(* CODESYS project YarnStorage.xml

Project tree, tasks and I/O mapping:
  visualisation YarnStorage
*)

// /YarnStorage
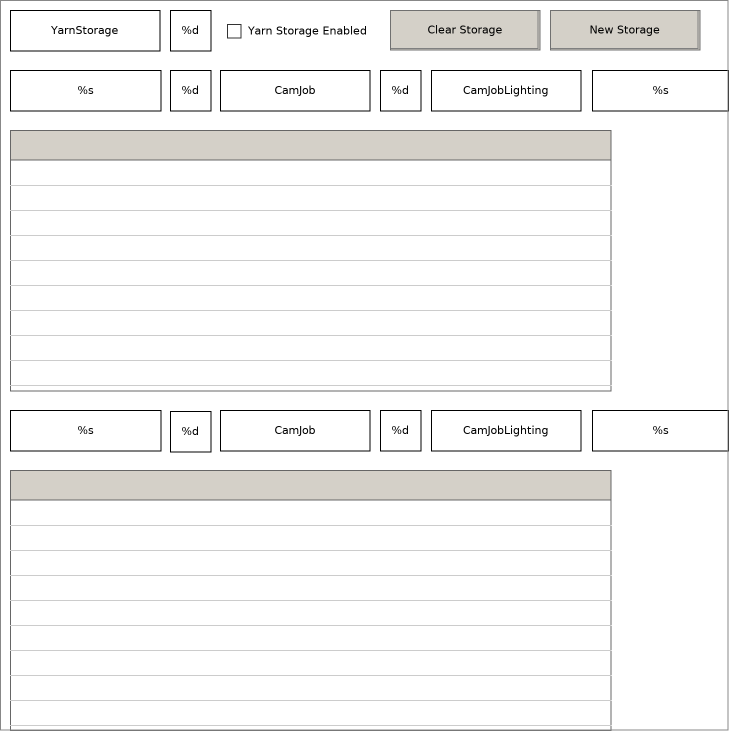
VISUALIZATION YarnStorage  // 729x731
    Rectangle (10,10 150x41), "YarnStorage"
    Rectangle (170,10 41x41), "%d", text variable: PRG_VisuTask_10ms._fbYarnStorageCtrl._iStorage
        OnMouseUp: write the text variable via Default
    Rectangle (10,70 151x41), "%s", text variable: PRG_VisuTask_10ms._fbYarnStorageCtrl._aState[1]
        OnMouseUp: write the text variable via Default
    Rectangle (10,410 151x41), "%s", text variable: PRG_VisuTask_10ms._fbYarnStorageCtrl._aState[2]
        OnMouseUp: write the text variable via Default
    Table (10,130 601x261), data array: PRG_VisuTask_10ms._fbYarnStorageCtrl._ascCoilPositionsBase
        p3854506369: PRG_VisuTask_10ms._fbYarnStorageCtrl._ascCoilPositionsBase[INDEX].posX
        p1892666644: PRG_VisuTask_10ms._fbYarnStorageCtrl._ascCoilPositionsBase[INDEX].posY
        p338671338: PRG_VisuTask_10ms._fbYarnStorageCtrl._ascCoilPositionsBase[INDEX].posZ
        p2170511999: PRG_VisuTask_10ms._fbYarnStorageCtrl._ascCoilPositionsBase[INDEX].posRX
        p3723444502: PRG_VisuTask_10ms._fbYarnStorageCtrl._ascCoilPositionsBase[INDEX].posRY
        p1218418051: PRG_VisuTask_10ms._fbYarnStorageCtrl._ascCoilPositionsBase[INDEX].posRZ
        p746581629: PRG_VisuTask_10ms._fbYarnStorageCtrl._ascCoilPositionsBase[INDEX].offsetX1
        p3104783080: PRG_VisuTask_10ms._fbYarnStorageCtrl._ascCoilPositionsBase[INDEX].offsetY1
        p2501879983: PRG_VisuTask_10ms._fbYarnStorageCtrl._ascCoilPositionsBase[INDEX].offsetZ1
        p7306298: PRG_VisuTask_10ms._fbYarnStorageCtrl._ascCoilPositionsBase[INDEX].offsetX2
        p1933151965: PRG_VisuTask_10ms._fbYarnStorageCtrl._ascCoilPositionsBase[INDEX].offsetY2
        p3863566920: PRG_VisuTask_10ms._fbYarnStorageCtrl._ascCoilPositionsBase[INDEX].offsetZ2
        p2192122294: PRG_VisuTask_10ms._fbYarnStorageCtrl._ascCoilPositionsBase[INDEX].offsetX3
        p400160035: PRG_VisuTask_10ms._fbYarnStorageCtrl._ascCoilPositionsBase[INDEX].offsetY3
        p1265227338: PRG_VisuTask_10ms._fbYarnStorageCtrl._ascCoilPositionsBase[INDEX].offsetZ3
        p3726181087: PRG_VisuTask_10ms._fbYarnStorageCtrl._ascCoilPositionsBase[INDEX].offsetX4
        p3136911649: PRG_VisuTask_10ms._fbYarnStorageCtrl._ascCoilPositionsBase[INDEX].offsetY4
        p797552052: PRG_VisuTask_10ms._fbYarnStorageCtrl._ascCoilPositionsBase[INDEX].offsetZ4
        p60375027: PRG_VisuTask_10ms._fbYarnStorageCtrl._ascCoilPositionsBase[INDEX].offsetX5
        p2531912550: PRG_VisuTask_10ms._fbYarnStorageCtrl._ascCoilPositionsBase[INDEX].offsetY5
        p693678525: PRG_VisuTask_10ms._fbYarnStorageCtrl._ascCoilPositionsBase[INDEX].offsetZ5
        p3156763944: PRG_VisuTask_10ms._fbYarnStorageCtrl._ascCoilPositionsBase[INDEX].offsetX6
        p3636993750: PRG_VisuTask_10ms._fbYarnStorageCtrl._ascCoilPositionsBase[INDEX].offsetY6
        p1303956035: PRG_VisuTask_10ms._fbYarnStorageCtrl._ascCoilPositionsBase[INDEX].offsetZ6
        p285796650: PRG_VisuTask_10ms._fbYarnStorageCtrl._ascCoilPositionsBase[INDEX].offsetX7
        p2222472639: PRG_VisuTask_10ms._fbYarnStorageCtrl._ascCoilPositionsBase[INDEX].offsetY7
        p3768075841: PRG_VisuTask_10ms._fbYarnStorageCtrl._ascCoilPositionsBase[INDEX].offsetZ7
        p1978176212: PRG_VisuTask_10ms._fbYarnStorageCtrl._ascCoilPositionsBase[INDEX].offsetX8
        p1509425299: PRG_VisuTask_10ms._fbYarnStorageCtrl._ascCoilPositionsBase[INDEX].offsetY8
        p3431519238: PRG_VisuTask_10ms._fbYarnStorageCtrl._ascCoilPositionsBase[INDEX].offsetZ8
        p2846402210: PRG_VisuTask_10ms._fbYarnStorageCtrl._ascCoilPositionsBase[INDEX].offsetX9
        p1020817975: PRG_VisuTask_10ms._fbYarnStorageCtrl._ascCoilPositionsBase[INDEX].offsetY9
        p1480067529: PRG_VisuTask_10ms._fbYarnStorageCtrl._ascCoilPositionsBase[INDEX].offsetZ9
        p2232123230: Pos X
        p511219082: Pos Y
        p1014161805: GVL_Constant.cMaxNbrCoilPositions - 0 + 1
    Table (10,470 601x261), data array: PRG_VisuTask_10ms._fbYarnStorageCtrl._ascCoilPositionsInverted
        p3854506369: PRG_VisuTask_10ms._fbYarnStorageCtrl._ascCoilPositionsInverted[INDEX].posX
        p1892666644: PRG_VisuTask_10ms._fbYarnStorageCtrl._ascCoilPositionsInverted[INDEX].posY
        p338671338: PRG_VisuTask_10ms._fbYarnStorageCtrl._ascCoilPositionsInverted[INDEX].posZ
        p2170511999: PRG_VisuTask_10ms._fbYarnStorageCtrl._ascCoilPositionsInverted[INDEX].posRX
        p3723444502: PRG_VisuTask_10ms._fbYarnStorageCtrl._ascCoilPositionsInverted[INDEX].posRY
        p1218418051: PRG_VisuTask_10ms._fbYarnStorageCtrl._ascCoilPositionsInverted[INDEX].posRZ
        p746581629: PRG_VisuTask_10ms._fbYarnStorageCtrl._ascCoilPositionsInverted[INDEX].offsetX1
        p3104783080: PRG_VisuTask_10ms._fbYarnStorageCtrl._ascCoilPositionsInverted[INDEX].offsetY1
        p2501879983: PRG_VisuTask_10ms._fbYarnStorageCtrl._ascCoilPositionsInverted[INDEX].offsetZ1
        p7306298: PRG_VisuTask_10ms._fbYarnStorageCtrl._ascCoilPositionsInverted[INDEX].offsetX2
        p1933151965: PRG_VisuTask_10ms._fbYarnStorageCtrl._ascCoilPositionsInverted[INDEX].offsetY2
        p3863566920: PRG_VisuTask_10ms._fbYarnStorageCtrl._ascCoilPositionsInverted[INDEX].offsetZ2
        p2192122294: PRG_VisuTask_10ms._fbYarnStorageCtrl._ascCoilPositionsInverted[INDEX].offsetX3
        p400160035: PRG_VisuTask_10ms._fbYarnStorageCtrl._ascCoilPositionsInverted[INDEX].offsetY3
        p1265227338: PRG_VisuTask_10ms._fbYarnStorageCtrl._ascCoilPositionsInverted[INDEX].offsetZ3
        p3726181087: PRG_VisuTask_10ms._fbYarnStorageCtrl._ascCoilPositionsInverted[INDEX].offsetX4
        p3136911649: PRG_VisuTask_10ms._fbYarnStorageCtrl._ascCoilPositionsInverted[INDEX].offsetY4
        p797552052: PRG_VisuTask_10ms._fbYarnStorageCtrl._ascCoilPositionsInverted[INDEX].offsetZ4
        p60375027: PRG_VisuTask_10ms._fbYarnStorageCtrl._ascCoilPositionsInverted[INDEX].offsetX5
        p2531912550: PRG_VisuTask_10ms._fbYarnStorageCtrl._ascCoilPositionsInverted[INDEX].offsetY5
        p693678525: PRG_VisuTask_10ms._fbYarnStorageCtrl._ascCoilPositionsInverted[INDEX].offsetZ5
        p3156763944: PRG_VisuTask_10ms._fbYarnStorageCtrl._ascCoilPositionsInverted[INDEX].offsetX6
        p3636993750: PRG_VisuTask_10ms._fbYarnStorageCtrl._ascCoilPositionsInverted[INDEX].offsetY6
        p1303956035: PRG_VisuTask_10ms._fbYarnStorageCtrl._ascCoilPositionsInverted[INDEX].offsetZ6
        p285796650: PRG_VisuTask_10ms._fbYarnStorageCtrl._ascCoilPositionsInverted[INDEX].offsetX7
        p2222472639: PRG_VisuTask_10ms._fbYarnStorageCtrl._ascCoilPositionsInverted[INDEX].offsetY7
        p3768075841: PRG_VisuTask_10ms._fbYarnStorageCtrl._ascCoilPositionsInverted[INDEX].offsetZ7
        p1978176212: PRG_VisuTask_10ms._fbYarnStorageCtrl._ascCoilPositionsInverted[INDEX].offsetX8
        p1509425299: PRG_VisuTask_10ms._fbYarnStorageCtrl._ascCoilPositionsInverted[INDEX].offsetY8
        p3431519238: PRG_VisuTask_10ms._fbYarnStorageCtrl._ascCoilPositionsInverted[INDEX].offsetZ8
        p2846402210: PRG_VisuTask_10ms._fbYarnStorageCtrl._ascCoilPositionsInverted[INDEX].offsetX9
        p1020817975: PRG_VisuTask_10ms._fbYarnStorageCtrl._ascCoilPositionsInverted[INDEX].offsetY9
        p1480067529: PRG_VisuTask_10ms._fbYarnStorageCtrl._ascCoilPositionsInverted[INDEX].offsetZ9
        p2232123230: Pos X
        p511219082: Pos Y
        p1014161805: GVL_Constant.cMaxNbrCoilPositions - 0 + 1
    Rectangle (170,70 41x41), "%d", text variable: PRG_VisuTask_10ms._fbYarnStorageCtrl._NbrOfCoilsBase
        OnMouseUp: write the text variable via Default
    Rectangle (170,411 41x41), "%d", text variable: PRG_VisuTask_10ms._fbYarnStorageCtrl._NbrOfCoilsInverted
        OnMouseUp: write the text variable via Default
    Button (390,10 150x40), "Clear Storage", input disabled if: NOT PRG_VisuTask_10ms._fbManualCtrl.xManualMode
        tap PRG_VisuTask_10ms._fbYarnStorageCtrl._btnClearStorage.xbtn
    Checkbox (225,16 174x30), "Yarn Storage Enabled", variable: PersistentVars.scYarnStorages.ascYarnStorage[PRG_VisuTask_10ms._fbYarnStorageCtrl._iStorage].xEnabled
    Rectangle (431,70 150x41), "CamJobLighting"
    Rectangle (592,70 137x41), "%s", text variable: PRG_VisuTask_10ms._fbYarnStorageCtrl._CamLightingModeBase
        OnMouseUp: write the text variable via Default
    Rectangle (220,70 150x41), "CamJob"
    Rectangle (380,70 41x41), "%d", text variable: PRG_VisuTask_10ms._fbYarnStorageCtrl._CamJobBase
        OnMouseUp: write the text variable via Default
    Rectangle (220,410 150x41), "CamJob"
    Rectangle (380,410 41x41), "%d", text variable: PRG_VisuTask_10ms._fbYarnStorageCtrl._CamJobinverted
        OnMouseUp: write the text variable via Default
    Rectangle (431,410 150x41), "CamJobLighting"
    Rectangle (592,410 137x41), "%s", text variable: PRG_VisuTask_10ms._fbYarnStorageCtrl._CamLightingModeinverted
        OnMouseUp: write the text variable via Default
    Button (550,10 150x40), "New Storage"
        tap PRG_VisuTask_10ms._fbYarnStorageCtrl._btnNewPallet.xbtn
END_VISUALIZATION
